(* CODESYS project Alarms.export

Project tree, tasks and I/O mapping:
  visualisation Alarms
*)

// /Alarms
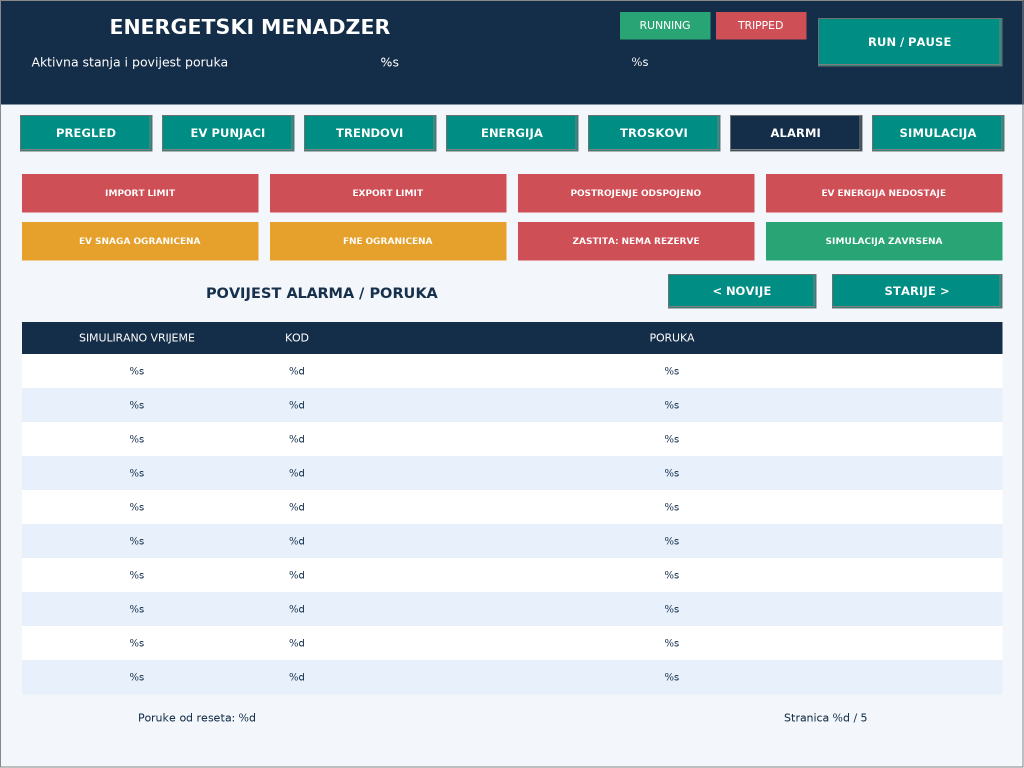
VISUALIZATION Alarms  // 1024x768
    Rectangle (0,0 1024x768)
    Rectangle (0,0 1024x104)
    Rectangle (20,10 460x34), "ENERGETSKI MENADZER"
    Rectangle (20,48 220x28), "Aktivna stanja i povijest poruka"
    Rectangle (260,49 260x26), "%s", text variable: Team_HMI.sDateTime
    Rectangle (530,49 220x26), "%s", text variable: Team_HMI.sPriceMode
    Button (818,18 184x48), "RUN / PAUSE"
        toggle SimCtrl.run
    Rectangle (620,12 90x27), "PAUSED", invisible if: SimCtrl.run
    Rectangle (620,12 90x27), "RUNNING", invisible if: NOT SimCtrl.run
    Rectangle (716,12 90x27), "TRIPPED", invisible if: NOT SimCtrl.tripped
    Button (20,115 132x36), "PREGLED"
        OnMouseClick:  Assign=Overview, Type=Assignment
    Button (162,115 132x36), "EV PUNJACI"
        OnMouseClick:  Assign=EVs, Type=Assignment
    Button (304,115 132x36), "TRENDOVI"
        OnMouseClick:  Assign=Trends, Type=Assignment
    Button (446,115 132x36), "ENERGIJA"
        OnMouseClick:  Assign=Energy, Type=Assignment
    Button (588,115 132x36), "TROSKOVI"
        OnMouseClick:  Assign=Costs, Type=Assignment
    Button (730,115 132x36), "ALARMI"
        OnMouseClick:  Assign=Alarms, Type=Assignment
    Button (872,115 132x36), "SIMULACIJA"
        OnMouseClick:  Assign=Controls, Type=Assignment
    Rectangle (22,174 236x38), "IMPORT LIMIT"
    Rectangle (22,174 236x38), "IMPORT LIMIT", invisible if: NOT Team_HMI.xAlmImport
    Rectangle (270,174 236x38), "EXPORT LIMIT"
    Rectangle (270,174 236x38), "EXPORT LIMIT", invisible if: NOT Team_HMI.xAlmExport
    Rectangle (518,174 236x38), "POSTROJENJE ODSPOJENO"
    Rectangle (518,174 236x38), "POSTROJENJE ODSPOJENO", invisible if: NOT Team_HMI.xAlmTripped
    Rectangle (766,174 236x38), "EV ENERGIJA NEDOSTAJE"
    Rectangle (766,174 236x38), "EV ENERGIJA NEDOSTAJE", invisible if: NOT Team_HMI.xAlmEvUnmet
    Rectangle (22,222 236x38), "EV SNAGA OGRANICENA"
    Rectangle (22,222 236x38), "EV SNAGA OGRANICENA", invisible if: NOT Team_HMI.xAlmGuardEv
    Rectangle (270,222 236x38), "FNE OGRANICENA"
    Rectangle (270,222 236x38), "FNE OGRANICENA", invisible if: NOT Team_HMI.xAlmGuardCurt
    Rectangle (518,222 236x38), "ZASTITA: NEMA REZERVE"
    Rectangle (518,222 236x38), "ZASTITA: NEMA REZERVE", invisible if: NOT Team_HMI.xAlmGuardFail
    Rectangle (766,222 236x38), "SIMULACIJA ZAVRSENA"
    Rectangle (766,222 236x38), "SIMULACIJA ZAVRSENA", invisible if: NOT Team_HMI.xAlmFinished
    Rectangle (22,278 600x30), "POVIJEST ALARMA / PORUKA"
    Button (668,274 148x34), "< NOVIJE"
        OnMouseClick: execute { Team_Visu.iAlarmPage := MAX(0, Team_Visu.iAlarmPage - 1); }
    Button (832,274 170x34), "STARIJE >"
        OnMouseClick: execute { Team_Visu.iAlarmPage := MIN(4, Team_Visu.iAlarmPage + 1); }
    Rectangle (22,322 230x32), "SIMULIRANO VRIJEME"
    Rectangle (252,322 90x32), "KOD"
    Rectangle (342,322 660x32), "PORUKA"
    Rectangle (22,354 230x34), "%s", text variable: Team_HMI.aAlarmHist[Team_Visu.iAlarmPage * 10 + 0].sStamp
    Rectangle (252,354 90x34), "%d", text variable: Team_HMI.aAlarmHist[Team_Visu.iAlarmPage * 10 + 0].iCode
    Rectangle (342,354 660x34), "%s", text variable: Team_HMI.aAlarmHist[Team_Visu.iAlarmPage * 10 + 0].sText
    Rectangle (22,388 230x34), "%s", text variable: Team_HMI.aAlarmHist[Team_Visu.iAlarmPage * 10 + 1].sStamp
    Rectangle (252,388 90x34), "%d", text variable: Team_HMI.aAlarmHist[Team_Visu.iAlarmPage * 10 + 1].iCode
    Rectangle (342,388 660x34), "%s", text variable: Team_HMI.aAlarmHist[Team_Visu.iAlarmPage * 10 + 1].sText
    Rectangle (22,422 230x34), "%s", text variable: Team_HMI.aAlarmHist[Team_Visu.iAlarmPage * 10 + 2].sStamp
    Rectangle (252,422 90x34), "%d", text variable: Team_HMI.aAlarmHist[Team_Visu.iAlarmPage * 10 + 2].iCode
    Rectangle (342,422 660x34), "%s", text variable: Team_HMI.aAlarmHist[Team_Visu.iAlarmPage * 10 + 2].sText
    Rectangle (22,456 230x34), "%s", text variable: Team_HMI.aAlarmHist[Team_Visu.iAlarmPage * 10 + 3].sStamp
    Rectangle (252,456 90x34), "%d", text variable: Team_HMI.aAlarmHist[Team_Visu.iAlarmPage * 10 + 3].iCode
    Rectangle (342,456 660x34), "%s", text variable: Team_HMI.aAlarmHist[Team_Visu.iAlarmPage * 10 + 3].sText
    Rectangle (22,490 230x34), "%s", text variable: Team_HMI.aAlarmHist[Team_Visu.iAlarmPage * 10 + 4].sStamp
    Rectangle (252,490 90x34), "%d", text variable: Team_HMI.aAlarmHist[Team_Visu.iAlarmPage * 10 + 4].iCode
    Rectangle (342,490 660x34), "%s", text variable: Team_HMI.aAlarmHist[Team_Visu.iAlarmPage * 10 + 4].sText
    Rectangle (22,524 230x34), "%s", text variable: Team_HMI.aAlarmHist[Team_Visu.iAlarmPage * 10 + 5].sStamp
    Rectangle (252,524 90x34), "%d", text variable: Team_HMI.aAlarmHist[Team_Visu.iAlarmPage * 10 + 5].iCode
    Rectangle (342,524 660x34), "%s", text variable: Team_HMI.aAlarmHist[Team_Visu.iAlarmPage * 10 + 5].sText
    Rectangle (22,558 230x34), "%s", text variable: Team_HMI.aAlarmHist[Team_Visu.iAlarmPage * 10 + 6].sStamp
    Rectangle (252,558 90x34), "%d", text variable: Team_HMI.aAlarmHist[Team_Visu.iAlarmPage * 10 + 6].iCode
    Rectangle (342,558 660x34), "%s", text variable: Team_HMI.aAlarmHist[Team_Visu.iAlarmPage * 10 + 6].sText
    Rectangle (22,592 230x34), "%s", text variable: Team_HMI.aAlarmHist[Team_Visu.iAlarmPage * 10 + 7].sStamp
    Rectangle (252,592 90x34), "%d", text variable: Team_HMI.aAlarmHist[Team_Visu.iAlarmPage * 10 + 7].iCode
    Rectangle (342,592 660x34), "%s", text variable: Team_HMI.aAlarmHist[Team_Visu.iAlarmPage * 10 + 7].sText
    Rectangle (22,626 230x34), "%s", text variable: Team_HMI.aAlarmHist[Team_Visu.iAlarmPage * 10 + 8].sStamp
    Rectangle (252,626 90x34), "%d", text variable: Team_HMI.aAlarmHist[Team_Visu.iAlarmPage * 10 + 8].iCode
    Rectangle (342,626 660x34), "%s", text variable: Team_HMI.aAlarmHist[Team_Visu.iAlarmPage * 10 + 8].sText
    Rectangle (22,660 230x34), "%s", text variable: Team_HMI.aAlarmHist[Team_Visu.iAlarmPage * 10 + 9].sStamp
    Rectangle (252,660 90x34), "%d", text variable: Team_HMI.aAlarmHist[Team_Visu.iAlarmPage * 10 + 9].iCode
    Rectangle (342,660 660x34), "%s", text variable: Team_HMI.aAlarmHist[Team_Visu.iAlarmPage * 10 + 9].sText
    Rectangle (22,704 350x28), "Poruke od reseta: %d", text variable: Team_HMI.nAlarms
    Rectangle (650,704 352x28), "Stranica %d / 5", text variable: Team_Visu.iAlarmPage + 1
END_VISUALIZATION
